Fanuc KAREL source: ko00089.KL

-- PROVISIONAL review KL for V770-1; original PC SHA256 554143e989866ccd5865345739a24e2d0bad2e878ae028afa3a6b00284c5bcea
-- Incomplete behavior may be omitted. Consult companion uncertainty JSON. Do not deploy.
PROGRAM KO00089
%NOLOCKGROUP
BEGIN
  -- UNRESOLVED_PC offsets 5-12; opcodes 9D,23
  -- UNRESOLVED_PC offsets 17-69; opcodes 27,27,49,7E,AD,27,49,7E,AD,22,31,7E,4A
  -- UNRESOLVED_PC offsets 74-78; opcodes 7F
END KO00089
